Fanuc KAREL source: kb00020.compact.KL

PROGRAM KB00020
%STACKSIZE=65535
%PRIORITY=65535
%NOLOCKGROUP
VAR
P1 : INTEGER
RESULT : STRING[80]
BEGIN
P1=1
RESULT=CHR(P1)
END KB00020
